(*
SPDX-FileCopyrightText: © 2026 Oleksandr Tiutyk <trofimich@gmail.com>
SPDX-License-Identifier: MIT
License: https://opensource.org/license/mit
*)

(*!
<summary>Provides fluent assertions on a copied DATE value.</summary>
<description>
Copies actual into persistent instance storage before the entry method returns; literals and expression
results therefore remain valid throughout the immediate chain. Owns no heap allocation or pointed-to resource.
The message prefixes every failure until the next preparation. Finish one chain before starting another on
the owning Assertions provider. Use only from the owning test callback on one task, without reentry.
Obtain this context from the owning provider; direct unprepared use is unsupported.
Expected arguments use the declared IEC type; ordinary compiler conversions happen before comparison.
This context does not depend on another assertion context.
Object metadata is available before preparation; inherited equality compares instance identity.
</description>
*)

{attribute 'no_explicit_call' := 'do not call this function block directly'}
FUNCTION_BLOCK DateAssertionContext EXTENDS TOF_Core.Object
VAR_STAT
	{attribute 'hide'}
	_ClassName : STRING := __POUNAME();
END_VAR
VAR
	_Actual : DATE;
	_TestCase : ITestCase;
	_Message : WSTRING(255);
END_VAR

(*!
<summary>Provides the implementation class name.</summary>
<description>
Borrowed read-only reference to compiler-initialized storage, valid throughout the instance lifetime.
Do not modify the returned reference; no ownership is transferred.
</description>
*)
{attribute 'monitoring' := 'call'}
PROPERTY ClassName : REFERENCE TO STRING
GET
ClassName REF= _ClassName;
END_GET
END_PROPERTY

(*!
<summary>Asserts that the actual value is strictly greater than expected.</summary>
<description>
Records failure without interrupting the callback; preserves the message for the rest of the chain.
</description>
<param name="expected">Expected value converted by the compiler to DATE.</param>
*)
METHOD FINAL IsGreaterThan : REFERENCE TO DateAssertionContext
VAR_INPUT
	expected : DATE;
END_VAR
IF _Actual <= expected THEN
	failComparison(
		expected := expected,
		expectation := "Expected value > "
	);
END_IF

IsGreaterThan REF= THIS^;
END_METHOD

(*!
<summary>Asserts that the actual value meets the inclusive lower boundary.</summary>
<description>
Records failure without interrupting the callback; preserves the message for the rest of the chain.
</description>
<param name="expected">Expected value converted by the compiler to DATE.</param>
*)
METHOD FINAL IsGreaterThanOrEquals : REFERENCE TO DateAssertionContext
VAR_INPUT
	expected : DATE;
END_VAR
IF _Actual < expected THEN
	failComparison(
		expected := expected,
		expectation := "Expected value >= "
	);
END_IF

IsGreaterThanOrEquals REF= THIS^;
END_METHOD

(*!
<summary>Asserts that the actual value is strictly less than expected.</summary>
<description>
Records failure without interrupting the callback; preserves the message for the rest of the chain.
</description>
<param name="expected">Expected value converted by the compiler to DATE.</param>
*)
METHOD FINAL IsLessThan : REFERENCE TO DateAssertionContext
VAR_INPUT
	expected : DATE;
END_VAR
IF _Actual >= expected THEN
	failComparison(
		expected := expected,
		expectation := "Expected value < "
	);
END_IF

IsLessThan REF= THIS^;
END_METHOD

(*!
<summary>Asserts that the actual value meets the inclusive upper boundary.</summary>
<description>
Records failure without interrupting the callback; preserves the message for the rest of the chain.
</description>
<param name="expected">Expected value converted by the compiler to DATE.</param>
*)
METHOD FINAL IsLessThanOrEquals : REFERENCE TO DateAssertionContext
VAR_INPUT
	expected : DATE;
END_VAR
IF _Actual > expected THEN
	failComparison(
		expected := expected,
		expectation := "Expected value <= "
	);
END_IF

IsLessThanOrEquals REF= THIS^;
END_METHOD

(*!
<summary>Provides the library namespace.</summary>
<description>
Borrowed read-only reference to the compiler-initialized namespace, valid throughout the instance lifetime.
Do not modify the returned reference; no ownership is transferred.
</description>
*)
{attribute 'monitoring' := 'call'}
PROPERTY NamespaceName : REFERENCE TO STRING
GET
NamespaceName REF= CurrentNamespace.Name;
END_GET
END_PROPERTY

(*!
<summary>Asserts inequality with the expected value.</summary>
<description>
Records failure without interrupting the callback; preserves the message for the rest of the chain.
</description>
<param name="expected">Expected value converted by the compiler to DATE.</param>
*)
METHOD FINAL NotToBe : REFERENCE TO DateAssertionContext
VAR_INPUT
	expected : DATE;
END_VAR
IF _Actual = expected THEN
	failComparison(
		expected := expected,
		expectation := "Expected value not to be: "
	);
END_IF

NotToBe REF= THIS^;
END_METHOD

(*!
<summary>Copies the actual operand and replaces the chain-wide message.</summary>
<description>
Called by the owning Assertions provider after it verifies the running test case.
No pointer to this method's input storage is retained. The receiver is borrowed until the next preparation;
the owning provider keeps it alive throughout the immediate chain.
</description>
<param name="actual">Value copied into this context.</param>
<param name="testCase">Borrowed failure receiver for the immediate chain.</param>
<param name="message">Copied diagnostic prefix, including empty to clear the previous prefix.</param>
*)
METHOD INTERNAL FINAL Prepare
VAR_INPUT
	actual : DATE;
	testCase : ITestCase;
END_VAR
VAR_IN_OUT CONSTANT
	message : WSTRING(255);
END_VAR
_Actual := actual;
_TestCase := testCase;
_Message := message;
END_METHOD

(*!
<summary>Reports the byte size of this concrete instance.</summary>
<description>
Includes inline fields and nested instances, but excludes separately allocated payloads.
Obtaining the size does not transfer ownership or validate an arbitrary address.
</description>
*)
{attribute 'monitoring' := 'call'}
PROPERTY SelfSize : ULINT
GET
SelfSize := XSIZEOF(THIS^);
END_GET
END_PROPERTY

(*!
<summary>Asserts equality with the expected value.</summary>
<description>
Records failure without interrupting the callback; preserves the message for the rest of the chain.
</description>
<param name="expected">Expected value converted by the compiler to DATE.</param>
*)
METHOD FINAL ToBe : REFERENCE TO DateAssertionContext
VAR_INPUT
	expected : DATE;
END_VAR
IF _Actual <> expected THEN
	failComparison(
		expected := expected,
		expectation := "Expected: "
	);
END_IF

ToBe REF= THIS^;
END_METHOD

(*!
<summary>Formats a failed typed predicate and reports it with the chain message.</summary>
<description>
Does not change operands or chain state. The receiver retains its first failure. Reporting exceptions
propagate to the enclosing test callback handler; an unprepared receiver is a configuration error.
</description>
<param name="expected">Typed expected operand used only for this diagnostic.</param>
<param name="expectation">Prefix identifying the failed predicate.</param>
*)
METHOD PRIVATE failComparison
VAR_INPUT
	expected : DATE;
	expectation : WSTRING(40);
END_VAR
VAR
	actualText : WSTRING(255);
	expectedText : WSTRING(255);
	diagnostic : TOF_Core.ERROR_MESSAGE;
END_VAR
actualText := TO_WSTRING(_Actual);
expectedText := TO_WSTRING(expected);

diagnostic := TOF_Core.WideStrings.Concat255(
	expectation,
	expectedText,
	", but was: ",
	actualText
);

TestServices.ReportAssertionFailure(
	testCase := _TestCase,
	message := _Message,
	sourceClassName := ClassName,
	defaultMessage := diagnostic
);
END_METHOD

END_FUNCTION_BLOCK

(* stored: Version 1.1.0.1
   POU DateAssertionContext: Id {e34d68b4-69aa-492f-b2a1-80eb8e630183}, SpecialFunc None
   Folder Service methods: Id {62d4da3b-efda-4275-ab09-ebfaf34af50c}
   Property ClassName: Id {e969be37-7933-4148-b15e-424831f13bc3}
   Get Get: Id {8a964911-9a1d-40fb-a302-bd294aa327ab}
   Method IsGreaterThan: Id {593f3be7-9e4f-4faa-9961-78992b1e798c}
   Method IsGreaterThanOrEquals: Id {48b215af-e91e-4f16-b2b1-54f06a51e8da}
   Method IsLessThan: Id {1bc67dbb-cdbb-40f8-b576-b6d7b51b5cc9}
   Method IsLessThanOrEquals: Id {45897868-35be-418d-b90b-49596184133b}
   Property NamespaceName: Id {30d5a921-f1e1-404d-ba16-214fc8be943b}
   Get Get: Id {8568e411-88cf-4283-a27f-5a4a5a511ac2}
   Method NotToBe: Id {767b7ab8-a6e3-47f0-814f-4d2e6cdd1061}
   Method Prepare: Id {3c935b06-7374-4c6b-a1e3-79e92078bb77}
   Property SelfSize: Id {5ce103ce-246c-40c5-aed7-8c574a267c59}
   Get Get: Id {483c7dc1-d1ee-4d1a-aa35-aa8a67edd930}
   Method ToBe: Id {3bd97314-45b2-4a1b-8d73-8c280ef217e9}
   Method failComparison: Id {3c5dc580-101f-46dd-8488-2cbdc64ac148} *)
